(* IEC 61131-3 sources: ayran-mini-fabrika/plc/build (part 2) *)

  CASE STP OF
    0:  (* idle *)
      WANT := WORD#0;
      PUMP_REQ := FALSE;
      IF NOT WAIT_START AND (ALARMS AND ALARM_MASK) = WORD#0 THEN
        IF CIP_REQ THEN
          CIP_REQ := FALSE;
          STP := 40;
        ELSIF REQ AND NOT CIP_DUE AND NOT DI_T1_LOW THEN
          BATCH := 0;
          IF LINE_PRODUCT THEN STP := 10; ELSE STP := 20; END_IF;
        END_IF;
      END_IF;

    20: (* fill the line with product: first liquid to the drain *)
      WANT := WORD#16#0022;            (* V_PROD + V_DRAIN *)
      PUMP_REQ := TRUE;
      IF T_INWIN.Q THEN
        LINE_PRODUCT := TRUE;
        STP := 10;                     (* the route manager stops the pump and changes the route *)
      ELSIF STEP_SCANS > 2250 THEN
        ALARMS := ALARMS OR WORD#16#0200;   (* product conductivity not detected within 45 s *)
      END_IF;

    10: (* transfer to the filling tank *)
      WANT := WORD#16#0012;            (* V_PROD + V_FILL *)
      PUMP_REQ := TRUE;
      IF T_FOREIGN.Q THEN
        LINE_PRODUCT := FALSE;
        ALARMS := ALARMS OR WORD#16#0004;
      ELSIF NOT REQ OR DI_T1_LOW OR SINCE >= CIP_LIMIT OR CIP_REQ THEN
        STP := 0;
      END_IF;

    40: (* CIP preparation: empty route for the line, prove all valves closed *)
      WANT := WORD#0;
      PUMP_REQ := FALSE;
      LINE_PRODUCT := FALSE;
      CAUSTIC_IN := FALSE;
      CIP_SCANS := 0;
      MIN_T := 32000;
      MIN_F := 32000;
      FINAL_COND := 0;
      IF IW_CIP_LVL < CIP_LVL_MIN THEN
        ALARMS := ALARMS OR WORD#16#0100;
      ELSIF RSTATE = 0 AND ROUTE_OK THEN
        STP := 41;
      END_IF;

    41: (* wait for the caustic temperature *)
      WANT := WORD#0;
      PUMP_REQ := FALSE;
      IF IW_CIP_T >= CAUSTIC_SP - 50 THEN
        STP := 42;
      ELSIF STEP_TO THEN
        ALARMS := ALARMS OR WORD#16#0080;
      END_IF;

    42: (* pre-rinse: water to the drain *)
      WANT := WORD#16#0024;            (* V_WATER + V_DRAIN *)
      PUMP_REQ := TRUE;
      IF VOL >= RINSE_KG THEN
        WATER_REF := IW_COND;           (* conductivity of the inlet water: the criterion for the final rinse *)
        STP := 43;
      ELSIF STEP_TO THEN
        ALARMS := ALARMS OR WORD#16#0080;
      END_IF;

    43: (* caustic: first to the drain, to the caustic tank once caustic arrives (phase separation) *)
      PUMP_REQ := TRUE;
      IF NOT CAUSTIC_IN AND RSTATE = 0 AND IW_COND >= COND_CAUSTIC THEN CAUSTIC_IN := TRUE; END_IF;
      IF CAUSTIC_IN THEN
        WANT := WORD#16#0048;          (* V_CAUSTIC + V_CIPRET *)
      ELSE
        WANT := WORD#16#0028;          (* V_CAUSTIC + V_DRAIN *)
      END_IF;
      (* CIP record: the lowest values in the counted hold window *)
      IF HOLD_OK THEN
        IF IW_RET_T < MIN_T THEN MIN_T := IW_RET_T; END_IF;
        IF IW_FLOW < MIN_F THEN MIN_F := IW_FLOW; END_IF;
      ELSE
        MIN_T := 32000;
        MIN_F := 32000;
      END_IF;
      IF T_HOLD.Q THEN
        STP := 44;
      ELSIF STEP_TO THEN
        ALARMS := ALARMS OR WORD#16#0080;
      END_IF;

    44: (* final rinse: until no caustic is left *)
      WANT := WORD#16#0024;
      PUMP_REQ := TRUE;
      IF VOL >= RINSE_KG AND IW_COND <= WATER_REF + RINSE_MARGIN THEN
        FINAL_COND := IW_COND;
        STP := 45;
      ELSIF STEP_TO THEN
        ALARMS := ALARMS OR WORD#16#0080;
      END_IF;

    45: (* completed *)
      WANT := WORD#0;
      PUMP_REQ := FALSE;
      SINCE := 0;
      CIP_DUE := FALSE;
      ABORT_WARN := FALSE;
      CIP_RES := 1;
      CIP_DUR := CIP_SCANS / 50;
      STP := 0;
  END_CASE;
  IF STP >= 40 AND STP <= 44 AND CIP_SCANS < 30000 THEN CIP_SCANS := CIP_SCANS + 1; END_IF;
  IF CIP_RES = 2 OR CIP_RES = 3 THEN CIP_DUR := CIP_SCANS / 50; END_IF;

  (* =================== 4. Route manager =================== *)
  IF (ALARMS AND ALARM_MASK) <> WORD#0 THEN WANT := WORD#0; END_IF;
  IF WANT <> CUR AND RSTATE = 0 THEN RSTATE := 1; END_IF;
  T_ROUTE(IN := RSTATE = 1, PT := T#3s);
  T_STROKE(IN := RSTATE = 2, PT := T#1s);
  IF RSTATE = 1 THEN
    VALVES := CUR AND WANT;            (* close the ones not in the new route *)
    IF ((NOT WANT) AND WORD#16#007E AND (NOT CLOSED)) = WORD#0 THEN
      RSTATE := 2;
    ELSIF T_ROUTE.Q THEN
      ALARMS := ALARMS OR WORD#16#0008;
      RSTATE := 0;
      CUR := CUR AND WANT;
    END_IF;
  ELSIF RSTATE = 2 THEN
    VALVES := WANT;
    IF T_STROKE.Q THEN CUR := WANT; RSTATE := 0; END_IF;
  ELSE
    VALVES := CUR;
  END_IF;

  Q_P1 := PUMP_REQ AND RSTATE = 0 AND CUR = WANT AND CUR <> WORD#0 AND ROUTE_OK
          AND (ALARMS AND ALARM_MASK) = WORD#0;

  (* caustic tank thermostat (+/- 2 C), level and over-temperature interlock *)
  IF NOT ESTOP_OK OR IW_CIP_LVL < CIP_LVL_MIN OR IW_CIP_T > CAUSTIC_MAX THEN
    Q_HEAT := FALSE;
  ELSIF IW_CIP_T < CAUSTIC_SP - 20 THEN
    Q_HEAT := TRUE;
  ELSIF IW_CIP_T > CAUSTIC_SP + 20 THEN
    Q_HEAT := FALSE;
  END_IF;

  (* =================== 5. Outputs =================== *)
  WARNS := WORD#0;
  IF DI_T1_LOW THEN WARNS := WARNS OR WORD#16#0400; END_IF;
  IF CIP_DUE THEN WARNS := WARNS OR WORD#16#0800; END_IF;
  IF ABORT_WARN THEN WARNS := WARNS OR WORD#16#1000; END_IF;

  QW_DO := VALVES AND WORD#16#007E;
  IF Q_P1 THEN QW_DO := QW_DO OR WORD#16#0001; END_IF;
  IF Q_HEAT THEN QW_DO := QW_DO OR WORD#16#0080; END_IF;
  IF STP >= 40 THEN QW_DO := QW_DO OR WORD#16#0100; END_IF;

  IF (ALARMS AND WORD#16#0001) <> WORD#0 THEN
    QW_STATE := 11;
  ELSIF (ALARMS AND ALARM_MASK) <> WORD#0 THEN
    QW_STATE := 10;
  ELSIF STP = 0 AND CIP_DUE THEN
    QW_STATE := 9;
  ELSIF STP = 0 THEN
    QW_STATE := 0;
  ELSIF (STP = 10 OR STP = 20) AND RSTATE <> 0 THEN
    QW_STATE := 3;
  ELSIF STP = 10 THEN
    QW_STATE := 1;
  ELSIF STP = 20 THEN
    QW_STATE := 2;
  ELSE
    QW_STATE := STP - 36;             (* 40..44 -> 4..8 *)
  END_IF;

  QW_ALARM    := ALARMS OR WARNS;
  QW_STEP_T   := STEP_SCANS / 50;
  QW_SINCE    := SINCE;
  QW_BATCH    := BATCH;
  QW_CIP_RES  := CIP_RES;
  IF MIN_T = 32000 THEN QW_CIP_MINT := 0; ELSE QW_CIP_MINT := MIN_T; END_IF;
  IF MIN_F = 32000 THEN QW_CIP_MINF := 0; ELSE QW_CIP_MINF := MIN_F; END_IF;
  QW_CIP_COND := FINAL_COND;
  QW_CIP_DUR  := CIP_DUR;
  TRANSFERRING := STP = 10 AND Q_P1;
  QW_STATUS := WORD#0;
  IF WAIT_START THEN QW_STATUS := WORD#16#0080; END_IF;
  IF WAIT_START OR NOT IO_READY THEN
    QW_DO := WORD#0;
    Q_HEAT := FALSE; Q_P1 := FALSE;
  END_IF;
END_FUNCTION_BLOCK

PROGRAM Fabrika
  VAR
    (* --- blok 0: Fabrika --- *)
    FAB_IW_DI        AT %IW100 : WORD;  (* Fabrika paneli girisleri (bit paketli) *)
    FAB_IW_MAPVER    AT %IW101 : INT;  (* Sinyal haritasi surumu *)
    FAB_IW_SIM_HB    AT %IW102 : INT;  (* Simulator kalp atisi (100 ms) *)
    FAB_QW_DO        AT %QW100 : WORD;  (* Fabrika cikislari (bit paketli) *)
    FAB_QW_PLC_HB    AT %QW101 : INT;  (* Proses PLC (ya da tek PLC) kalp atisi (her tarama) *)
    FAB_QW_STATE     AT %QW102 : INT;  (* Fabrika durumu *)
    FAB_QW_ALARM     AT %QW103 : WORD;  (* Fabrika alarm ozeti *)
    (* --- blok 1: Dolum-kapama --- *)
    DOL_IW_DI        AT %IW116 : WORD;  (* Dijital girisler (bit paketli) *)
    DOL_IW_FILL      AT %IW117 : INT;  (* Dolum terazisi (net) *)
    DOL_IW_TANK      AT %IW118 : INT;  (* Dolum tanki seviyesi *)
    DOL_IW_TEMP      AT %IW119 : INT;  (* Kapama kafasi sicakligi *)
    DOL_IW_CHECK     AT %IW120 : INT;  (* Kontrol tartisi (brut) *)
    DOL_QW_DO        AT %QW116 : WORD;  (* Dijital cikislar (bit paketli) *)
    DOL_QW_STATE     AT %QW117 : INT;  (* Makine modu *)
    DOL_QW_ALARM     AT %QW118 : WORD;  (* Alarm kelimesi *)
    DOL_QW_GOOD      AT %QW119 : INT;  (* Saglam bardak sayaci *)
    DOL_QW_REJECT    AT %QW120 : INT;  (* Red sayaci *)
    DOL_QW_STATUS    AT %QW121 : WORD;  (* Durum bitleri (bit 7: yeniden basladi, START bekliyor) *)
    (* --- blok 2: Tank ve transfer --- *)
    TNK_IW_DI        AT %IW132 : WORD;  (* Dijital girisler (bit paketli) *)
    TNK_IW_T1_LVL    AT %IW133 : INT;  (* Uretim tanki T1 seviyesi *)
    TNK_IW_FLOW      AT %IW134 : INT;  (* Debimetre FT1 *)
    TNK_IW_TOTAL     AT %IW135 : INT;  (* Debimetre toplayici (30000'de sifirlanir) *)
    TNK_IW_COND      AT %IW136 : INT;  (* Hat iletkenligi QT1 (25 ?C'ye duzeltilmis) *)
    TNK_IW_RET_T     AT %IW137 : INT;  (* Hat donus sicakligi TT1 *)
    TNK_IW_CIP_T     AT %IW138 : INT;  (* Kostik tanki sicakligi TT2 *)
    TNK_IW_CIP_LVL   AT %IW139 : INT;  (* Kostik tanki seviyesi *)
    TNK_QW_DO        AT %QW132 : WORD;  (* Dijital cikislar (bit paketli) *)
    TNK_QW_STATE     AT %QW133 : INT;  (* Istasyon durumu *)
    TNK_QW_ALARM     AT %QW134 : WORD;  (* Alarm kelimesi *)
    TNK_QW_STEP_T    AT %QW135 : INT;  (* Adim suresi *)
    TNK_QW_SINCE     AT %QW136 : INT;  (* Son CIP'ten beri aktarilan *)
    TNK_QW_BATCH     AT %QW137 : INT;  (* Bu aktarimda aktarilan *)
    TNK_QW_CIP_RES   AT %QW138 : INT;  (* Son CIP sonucu (0 yok, 1 basarili, 2 iptal, 3 basarisiz) *)
    TNK_QW_CIP_MINT  AT %QW139 : INT;  (* Son CIP: tutma sirasinda en dusuk donus sicakligi *)
    TNK_QW_CIP_MINF  AT %QW140 : INT;  (* Son CIP: tutma sirasinda en dusuk debi *)
    TNK_QW_CIP_COND  AT %QW141 : INT;  (* Son CIP: son durulama iletkenligi *)
    TNK_QW_CIP_DUR   AT %QW142 : INT;  (* Son CIP: toplam sure *)
    TNK_QW_STATUS    AT %QW143 : WORD;  (* Durum bitleri (bit 7: yeniden basladi, START bekliyor) *)
    (* --- blok 3: Shrink ve firin --- *)
    SHR_IW_DI        AT %IW148 : WORD;  (* Dijital girisler (bit paketli) *)
    SHR_IW_LANE      AT %IW149 : INT;  (* Seritteki bardak sayisi (bilesik sensor) *)
    SHR_IW_TEMP      AT %IW150 : INT;  (* Firin hava sicakligi *)
    SHR_IW_IN_CNT    AT %IW151 : INT;  (* Firin girisi paket sayaci (30000'de sifirlanir) *)
    SHR_IW_OUT_CNT   AT %IW152 : INT;  (* Firin cikisi paket sayaci *)
    SHR_IW_FILM      AT %IW153 : INT;  (* Film bobini kalan *)
    SHR_IW_PADS      AT %IW154 : INT;  (* Altlik magazini adedi *)
    SHR_IW_EXIT_CNT  AT %IW155 : INT;  (* Cikistan alinan paket sayaci *)
    SHR_IW_PLATE     AT %IW156 : WORD;  (* Plaka fotoselleri (bit 0: sira 1, bit 1: sira 2) *)
    SHR_IW_DIVERT    AT %IW157 : WORD;  (* Cikis ayirici: bit 0 paket var, 1 red konumu, 2 gecis konumu *)
    SHR_IW_REJECT_CNT AT %IW158 : INT;  (* Karantina kasasina ayrilan paket sayaci (30000 modul) *)
    SHR_QW_DO        AT %QW148 : WORD;  (* Dijital cikislar (bit paketli) *)
    SHR_QW_STATE     AT %QW149 : INT;  (* Istasyon durumu *)
    SHR_QW_ALARM     AT %QW150 : WORD;  (* Alarm kelimesi *)
    SHR_QW_STATUS    AT %QW151 : WORD;  (* Durum bitleri (PackML benzeri) *)
    SHR_QW_PACKS     AT %QW152 : INT;  (* Firina birakilan paket sayaci *)
    SHR_QW_INSIDE    AT %QW153 : INT;  (* Firin icindeki paket *)
    SHR_QW_SP        AT %QW154 : INT;  (* Gecerli firin ayar degeri *)
    SHR_QW_REJECT    AT %QW155 : INT;  (* Fotoselden dogrulanan karantina paket sayaci (30000 modul) *)
    SHR_QW_GOOD      AT %QW156 : INT;  (* Iyi urun bandina gecirilen paket sayaci (30000 modul) *)
    SHR_QW_PLC_HB    AT %QW163 : INT;  (* Paketleme PLC kalp atisi (her tarama) *)
    (* --- blok 4: Paletleme --- *)
    PAL_IW_DI        AT %IW164 : WORD;  (* Hat ve guvenlik girisleri (bit paketli) *)
    PAL_IW_ROB_DI    AT %IW165 : WORD;  (* Robot kontrolcusu durum bitleri *)
    PAL_IW_ACK_SEQ   AT %IW166 : INT;  (* Robot: kabul edilen son is numarasi *)
    PAL_IW_RES_SEQ   AT %IW167 : INT;  (* Robot: biten son is numarasi *)
    PAL_IW_RES_CODE  AT %IW168 : INT;  (* Robot: son is sonucu (1 tamam, 10+ hata) *)
    PAL_IW_RES_SLOT  AT %IW169 : INT;  (* Robot: son isin slotu *)
    PAL_IW_TURNS     AT %IW170 : INT;  (* Strec sarma: bu cevrimdeki tur *)
    PAL_IW_PALLETS   AT %IW171 : INT;  (* Bos palet magazini adedi *)
    PAL_IW_SHEETS    AT %IW172 : INT;  (* Karton levha magazini adedi *)
    PAL_IW_PICKUP_CNT AT %IW173 : INT;  (* Alim noktasindan alinan palet sayaci *)
    PAL_IW_IL        AT %IW174 : WORD;  (* Istasyon el sikisma girisleri (AGV optik I/O) *)
    PAL_IW_RES_JOB   AT %IW175 : INT;  (* Robot: biten son isin tipi *)
    PAL_QW_DO        AT %QW164 : WORD;  (* Dijital cikislar (bit paketli) *)
    PAL_QW_JOB       AT %QW165 : INT;  (* Robot isi (1 al, 2 birak, 3 levha, 4 eve don) *)
    PAL_QW_SLOT      AT %QW166 : INT;  (* Robot slotu (birak: 1..18, levha: 0 alt / 1 ust) *)
    PAL_QW_SEQ       AT %QW167 : INT;  (* Robot is numarasi (degisince is baslar) *)
    PAL_QW_STATE     AT %QW168 : INT;  (* Istasyon durumu *)
    PAL_QW_ALARM     AT %QW169 : WORD;  (* Alarm kelimesi *)
    PAL_QW_STATUS    AT %QW170 : WORD;  (* Durum bitleri (PackML benzeri) *)
    PAL_QW_COUNT     AT %QW171 : INT;  (* Istifteki paletin paket sayisi (dogrulanmis) *)
    PAL_QW_DONE      AT %QW172 : INT;  (* Tamamlanan palet sayaci *)
    PAL_QW_PALLET_ID AT %QW173 : INT;  (* Istifteki paletin numarasi *)
    PAL_QW_WRAPPED   AT %QW174 : INT;  (* Streclenen palet sayaci *)
    (* --- blok 5: AGV transpalet --- *)
    AGV_IW_DI        AT %IW180 : WORD;  (* AGV durum bitleri *)
    AGV_IW_ACK_SEQ   AT %IW181 : INT;  (* AGV: kabul edilen son is *)
    AGV_IW_RES_SEQ   AT %IW182 : INT;  (* AGV: biten son is *)
    AGV_IW_RES_CODE  AT %IW183 : INT;  (* AGV: son is sonucu *)
    AGV_IW_BATTERY   AT %IW184 : INT;  (* Batarya *)
    AGV_IW_NODE      AT %IW185 : INT;  (* Bulundugu / gittigi dugum *)
    AGV_IW_LOAD_ID   AT %IW186 : INT;  (* Cataldaki paletin numarasi *)
    AGV_IW_DELIVERED AT %IW187 : INT;  (* Teslim edilen palet sayaci *)
    AGV_IW_IL        AT %IW188 : WORD;  (* Istasyon el sikisma girisleri (paletleme hucresinden kablo) *)
    AGV_QW_DO        AT %QW180 : WORD;  (* AGV ve istasyon izinleri (bit paketli) *)
    AGV_QW_ORDER     AT %QW181 : INT;  (* AGV isi (1 tasi D?depo, 2 yuku depoya birak, 3 sarj, 4 park) *)
    AGV_QW_SEQ       AT %QW182 : INT;  (* AGV is numarasi *)
    AGV_QW_STATE     AT %QW183 : INT;  (* AGV durumu *)
    AGV_QW_ALARM     AT %QW184 : WORD;  (* Alarm kelimesi *)
    AGV_QW_STATUS    AT %QW185 : WORD;  (* Durum bitleri *)
    AGV_QW_MOVES     AT %QW186 : INT;  (* Tamamlanan tasima sayaci *)
    AGV_QW_PLC_HB    AT %QW195 : INT;  (* Lojistik PLC kalp atisi (her tarama) *)
    (* --- blok 6: Otomatik depo --- *)
    ASRS_IW_DI       AT %IW196 : WORD;  (* Vinc, konveyor ve guvenlik bitleri *)
    ASRS_IW_ACK_SEQ  AT %IW197 : INT;  (* Vinc: kabul edilen son is *)
    ASRS_IW_RES_SEQ  AT %IW198 : INT;  (* Vinc: biten son is *)
    ASRS_IW_RES_CODE AT %IW199 : INT;  (* Vinc: son is sonucu *)
    ASRS_IW_RES_LOC  AT %IW200 : INT;  (* Vinc: son isin gozu *)
    ASRS_IW_RES_ID   AT %IW201 : INT;  (* Vinc: son iste okunan palet numarasi (0 bos) *)
    ASRS_IW_IN_ID    AT %IW202 : INT;  (* Giris okuyucusu: palet numarasi (0 okunamadi) *)
    ASRS_IW_FORK_ID  AT %IW203 : INT;  (* Vinc catalindaki palet numarasi *)
    ASRS_IW_TEMP     AT %IW204 : INT;  (* Depo sicakligi *)
    ASRS_IW_SHIP_REQ AT %IW205 : INT;  (* Sevkiyat siparisi sayaci (palet) *)
    ASRS_IW_SHIPPED  AT %IW206 : INT;  (* Kamyona yuklenen palet sayaci *)
    ASRS_QW_DO       AT %QW196 : WORD;  (* Dijital cikislar (bit paketli) *)
    ASRS_QW_JOB      AT %QW197 : INT;  (* Vinc isi (1 depola, 2 cikar, 3 eve don, 4 goz kontrolu) *)
    ASRS_QW_LOC      AT %QW198 : INT;  (* Goz numarasi (1..36) *)
    ASRS_QW_SEQ      AT %QW199 : INT;  (* Vinc is numarasi *)
    ASRS_QW_STATE    AT %QW200 : INT;  (* Depo durumu *)
    ASRS_QW_ALARM    AT %QW201 : WORD;  (* Alarm kelimesi *)
    ASRS_QW_STATUS   AT %QW202 : WORD;  (* Durum bitleri *)
    ASRS_QW_OCC_A    AT %QW203 : WORD;  (* PLC envanteri: dolu gozler 1-16 (bit) *)
    ASRS_QW_OCC_B    AT %QW204 : WORD;  (* PLC envanteri: dolu gozler 17-32 (bit) *)
    ASRS_QW_OCC_C    AT %QW205 : WORD;  (* PLC envanteri: dolu gozler 33-36 (bit) *)
    ASRS_QW_STOCK    AT %QW206 : INT;  (* Stoktaki palet *)
    ASRS_QW_UNKNOWN  AT %QW207 : INT;  (* Durumu belirsiz goz (kontrol bekliyor) *)
    ASRS_QW_STORED   AT %QW208 : INT;  (* Depolanan palet sayaci *)
    ASRS_QW_PICKED   AT %QW209 : INT;  (* Sevkiyata cikarilan palet sayaci *)
    ASRS_QW_NEXT_ID  AT %QW210 : INT;  (* Siradaki sevk paleti (FIFO, 0 yok) *)
    TNK_COMMISSION AT %MW0 : WORD;
    RET_MAGIC AT %MW32 : WORD;
    RET_MAPVER AT %MW33 : INT;
    PAL_COUNT AT %MW34 : INT;
    PAL_ID AT %MW35 : INT;
    PAL_DONE AT %MW36 : INT;
    PAL_WRAPPED AT %MW37 : INT;
    PAL_SHEETS AT %MW38 : WORD;
    PAL_LAST_SEQ AT %MW39 : INT;
    PAL_ACTIVE AT %MW40 : WORD;
    PAL_C_PHASE AT %MW41 : INT;
    PAL_UNDERWRAP AT %MW42 : WORD;
    RET_CHECK AT %MW43 : WORD;
  END_VAR

  VAR
    PB_START    : BOOL;   (* factory panel *)
    PB_STOP_OK  : BOOL;
    PB_ESTOP_OK : BOOL;
    PB_RESET    : BOOL;
    FIRST_SCAN  : BOOL := TRUE;
    RESTART     : BOOL;
    IO_READY    : BOOL;   (* first data arrived from the simulator with the correct version *)
    COMM_FAULT  : BOOL;
    SIM_HB_LAST : INT;
    PLC_HB      : INT;
    T_SIMHB     : TON;
    DOLUM       : FB_Dolum;
    TANK        : FB_Tank;
    SHRINK      : FB_Shrink;
    PALLET      : FB_Pallet;
    AGV         : FB_Agv;
    ASRS        : FB_Asrs;
  END_VAR

  (* =================== 1. Factory panel =================== *)
  PB_START    := (FAB_IW_DI AND WORD#16#0001) <> WORD#0;
  PB_STOP_OK  := (FAB_IW_DI AND WORD#16#0002) <> WORD#0;
  PB_ESTOP_OK := (FAB_IW_DI AND WORD#16#0004) <> WORD#0;
  PB_RESET    := (FAB_IW_DI AND WORD#16#0008) <> WORD#0;

  (* =================== 2. Communication watchdog =================== *)
  (* communication fault if the simulator heartbeat does not change for 2 s *)
  T_SIMHB(IN := (FAB_IW_SIM_HB = SIM_HB_LAST), PT := T#2s);
  SIM_HB_LAST := FAB_IW_SIM_HB;
  COMM_FAULT := T_SIMHB.Q;
  (* inputs are invalid until the first data arrives and the map version matches *)
  IF FAB_IW_SIM_HB <> 0 AND FAB_IW_MAPVER = 7 THEN IO_READY := TRUE; END_IF;

  RESTART := FIRST_SCAN AND IO_READY;
  IF RESTART THEN FIRST_SCAN := FALSE; END_IF;

  (* PLC heartbeat: the simulator watches it and switches off this PLC's outputs if the program stops *)
  PLC_HB := PLC_HB + 1;
  IF PLC_HB > 30000 THEN PLC_HB := 0; END_IF;

  (* =================== Fill-and-seal =================== *)
  DOLUM(START := PB_START, STOP_OK := PB_STOP_OK, ESTOP_OK := PB_ESTOP_OK, RESET := PB_RESET,
        RESTART := RESTART, IO_READY := IO_READY, COMM_FAULT := COMM_FAULT,
        IW_DI := DOL_IW_DI, IW_FILL := DOL_IW_FILL, IW_TANK := DOL_IW_TANK,
        IW_TEMP := DOL_IW_TEMP, IW_CHECK := DOL_IW_CHECK);
  DOL_QW_DO     := DOLUM.QW_DO;
  DOL_QW_STATE  := DOLUM.QW_STATE;
  DOL_QW_ALARM  := DOLUM.QW_ALARM;
  DOL_QW_GOOD   := DOLUM.QW_GOOD;
  DOL_QW_REJECT := DOLUM.QW_REJECT;
  DOL_QW_STATUS := DOLUM.QW_STATUS;

  (* handshake: the filling machine requests product, the tank station transfers it (same PLC) *)
  TANK(START := PB_START, TNK_COMMISSION := TNK_COMMISSION, ESTOP_OK := PB_ESTOP_OK, RESET := PB_RESET, RESTART := RESTART, IO_READY := IO_READY, COMM_FAULT := COMM_FAULT,
       REQ := DOLUM.PRODUCT_REQ,
       IW_DI := TNK_IW_DI, IW_T1_LVL := TNK_IW_T1_LVL, IW_FLOW := TNK_IW_FLOW, IW_TOTAL := TNK_IW_TOTAL,
       IW_COND := TNK_IW_COND, IW_RET_T := TNK_IW_RET_T, IW_CIP_T := TNK_IW_CIP_T, IW_CIP_LVL := TNK_IW_CIP_LVL);
  TNK_QW_DO       := TANK.QW_DO;
  TNK_QW_STATE    := TANK.QW_STATE;
  TNK_QW_ALARM    := TANK.QW_ALARM;
  TNK_QW_STEP_T   := TANK.QW_STEP_T;
  TNK_QW_SINCE    := TANK.QW_SINCE;
  TNK_QW_BATCH    := TANK.QW_BATCH;
  TNK_QW_CIP_RES  := TANK.QW_CIP_RES;
  TNK_QW_CIP_MINT := TANK.QW_CIP_MINT;
  TNK_QW_CIP_MINF := TANK.QW_CIP_MINF;
  TNK_QW_CIP_COND := TANK.QW_CIP_COND;
  TNK_QW_CIP_DUR  := TANK.QW_CIP_DUR;
  TNK_QW_STATUS := TANK.QW_STATUS;

  (* =================== Grouping, wrapping, shrink tunnel =================== *)
  (* contract: when the outfeed belt is full the filler already waits, and this station in turn
     releases no pack into the tunnel when its own outfeed is full *)
  SHRINK(START := PB_START, STOP_OK := PB_STOP_OK, ESTOP_OK := PB_ESTOP_OK, RESET := PB_RESET,
         RESTART := RESTART, IO_READY := IO_READY, COMM_FAULT := COMM_FAULT,
         IW_DI := SHR_IW_DI, IW_LANE := SHR_IW_LANE, IW_TEMP := SHR_IW_TEMP,
         IW_IN_CNT := SHR_IW_IN_CNT, IW_OUT_CNT := SHR_IW_OUT_CNT, IW_FILM := SHR_IW_FILM, IW_PADS := SHR_IW_PADS,
         IW_PLATE := SHR_IW_PLATE, IW_REJECT_CNT := SHR_IW_REJECT_CNT);
  SHR_QW_DO     := SHRINK.QW_DO;
  SHR_QW_STATE  := SHRINK.QW_STATE;
  SHR_QW_ALARM  := SHRINK.QW_ALARM;
  SHR_QW_STATUS := SHRINK.QW_STATUS;
  SHR_QW_PACKS  := SHRINK.QW_PACKS;
  SHR_QW_INSIDE := SHRINK.QW_INSIDE;
  SHR_QW_SP     := SHRINK.QW_SP;
  SHR_QW_REJECT := SHRINK.QW_REJECT;
  SHR_QW_GOOD := SHRINK.QW_GOOD;

  (* =================== Robotic palletizing =================== *)
  (* contract: if the robot does not take the pack at the pickup point, the tunnel outfeed fills up and
     the shrink tunnel accepts no new pack. The AGV's "forks outside the pickup point" signal is the
     optical signal the vehicle gives to the station: the station's own input (PAL_IW_IL bit 0); it
     does not pass through the logistics PLC. *)
  PALLET(START := PB_START, STOP_OK := PB_STOP_OK, ESTOP_OK := PB_ESTOP_OK, RESET := PB_RESET,
         RESTART := RESTART, IO_READY := IO_READY, COMM_FAULT := COMM_FAULT,
         IW_DI := PAL_IW_DI, IW_ROB_DI := PAL_IW_ROB_DI, IW_ACK_SEQ := PAL_IW_ACK_SEQ, IW_RES_SEQ := PAL_IW_RES_SEQ,
         IW_RES_JOB := PAL_IW_RES_JOB, IW_RES_CODE := PAL_IW_RES_CODE, IW_RES_SLOT := PAL_IW_RES_SLOT, IW_TURNS := PAL_IW_TURNS,
         IW_PALLETS := PAL_IW_PALLETS, IW_SHEETS := PAL_IW_SHEETS,
         AGV_CLEAR := (PAL_IW_IL AND WORD#16#0001) <> WORD#0,
         RET_MAGIC := RET_MAGIC, RET_MAPVER := RET_MAPVER, PAL_COUNT := PAL_COUNT, PAL_ID := PAL_ID,
         PAL_DONE := PAL_DONE, PAL_WRAPPED := PAL_WRAPPED, PAL_SHEETS := PAL_SHEETS,
         PAL_LAST_SEQ := PAL_LAST_SEQ, PAL_ACTIVE := PAL_ACTIVE, PAL_C_PHASE := PAL_C_PHASE,
         PAL_UNDERWRAP := PAL_UNDERWRAP, RET_CHECK := RET_CHECK);
  PAL_QW_DO        := PALLET.QW_DO;
  PAL_QW_JOB       := PALLET.QW_JOB;
  PAL_QW_SLOT      := PALLET.QW_SLOT;
  PAL_QW_SEQ       := PALLET.QW_SEQ;
  PAL_QW_STATE     := PALLET.QW_STATE;
  PAL_QW_ALARM     := PALLET.QW_ALARM;
  PAL_QW_STATUS    := PALLET.QW_STATUS;
  PAL_QW_COUNT     := PALLET.QW_COUNT;
  PAL_QW_DONE      := PALLET.QW_DONE;
  PAL_QW_PALLET_ID := PALLET.QW_PALLET_ID;
  PAL_QW_WRAPPED   := PALLET.QW_WRAPPED;

  (* =================== Automated cold store =================== *)
  (* the inbound conveyor runs only while the AGV forks are outside *)
  ASRS(START := PB_START, STOP_OK := PB_STOP_OK, ESTOP_OK := PB_ESTOP_OK, RESET := PB_RESET,
       RESTART := RESTART, IO_READY := IO_READY, COMM_FAULT := COMM_FAULT,
       IW_DI := ASRS_IW_DI, IW_ACK_SEQ := ASRS_IW_ACK_SEQ, IW_RES_SEQ := ASRS_IW_RES_SEQ,
       IW_RES_CODE := ASRS_IW_RES_CODE, IW_RES_LOC := ASRS_IW_RES_LOC, IW_RES_ID := ASRS_IW_RES_ID,
       IW_IN_ID := ASRS_IW_IN_ID, IW_FORK_ID := ASRS_IW_FORK_ID, IW_TEMP := ASRS_IW_TEMP,
       IW_SHIP_REQ := ASRS_IW_SHIP_REQ, AGV_CLEAR_IN := (AGV_IW_DI AND WORD#16#0080) <> WORD#0);
  ASRS_QW_DO      := ASRS.QW_DO;
  ASRS_QW_JOB     := ASRS.QW_JOB;
  ASRS_QW_LOC     := ASRS.QW_LOC;
  ASRS_QW_SEQ     := ASRS.QW_SEQ;
  ASRS_QW_STATE   := ASRS.QW_STATE;
  ASRS_QW_ALARM   := ASRS.QW_ALARM;
  ASRS_QW_STATUS  := ASRS.QW_STATUS;
  ASRS_QW_OCC_A   := ASRS.QW_OCC_A;
  ASRS_QW_OCC_B   := ASRS.QW_OCC_B;
  ASRS_QW_OCC_C   := ASRS.QW_OCC_C;
  ASRS_QW_STOCK   := ASRS.QW_STOCK;
  ASRS_QW_UNKNOWN := ASRS.QW_UNKNOWN;
  ASRS_QW_STORED  := ASRS.QW_STORED;
  ASRS_QW_PICKED  := ASRS.QW_PICKED;
  ASRS_QW_NEXT_ID := ASRS.QW_NEXT_ID;

  (* =================== AGV =================== *)
  (* moves pallets according to the palletizing cell and cold store permissions. "Pallet ready at the
     pickup point": in a single PLC, PALLET.PICKUP_RDY directly; in split mode, the wire from the
     packaging PLC's PAL_QW_DO bit 11 output (AGV_IW_IL bit 0). *)
  AGV(START := PB_START, STOP_OK := PB_STOP_OK, ESTOP_OK := PB_ESTOP_OK, RESET := PB_RESET,
      RESTART := RESTART, IO_READY := IO_READY, COMM_FAULT := COMM_FAULT,
      IW_DI := AGV_IW_DI, IW_ACK_SEQ := AGV_IW_ACK_SEQ, IW_RES_SEQ := AGV_IW_RES_SEQ,
      IW_RES_CODE := AGV_IW_RES_CODE, IW_BATTERY := AGV_IW_BATTERY,
      D_READY := PALLET.PICKUP_RDY, IN_READY := ASRS.IN_READY);
  AGV_QW_DO     := AGV.QW_DO;
  AGV_QW_ORDER  := AGV.QW_ORDER;
  AGV_QW_SEQ    := AGV.QW_SEQ;
  AGV_QW_STATE  := AGV.QW_STATE;
  AGV_QW_ALARM  := AGV.QW_ALARM;
  AGV_QW_STATUS := AGV.QW_STATUS;
  AGV_QW_MOVES  := AGV.QW_MOVES;

  (* =================== Factory summary (block 0) =================== *)
  FAB_QW_PLC_HB := PLC_HB;
  IF DOLUM.RUNNING THEN FAB_QW_DO := WORD#16#0001; ELSE FAB_QW_DO := WORD#0; END_IF;
  FAB_QW_STATE := DOLUM.QW_STATE;
  FAB_QW_ALARM := DOLUM.QW_ALARM OR TANK.QW_ALARM OR SHRINK.QW_ALARM OR PALLET.QW_ALARM OR ASRS.QW_ALARM OR AGV.QW_ALARM;

  SHR_QW_PLC_HB := PLC_HB;

  AGV_QW_PLC_HB := PLC_HB;
END_PROGRAM

CONFIGURATION Config0
  RESOURCE Res0 ON PLC
    TASK task0(INTERVAL := T#20ms, PRIORITY := 0);
    PROGRAM instance0 WITH task0 : Fabrika;
  END_RESOURCE
END_CONFIGURATION
